(* IEC 61131-3 sources: plc-vscode/tests/st/all/trust-platform/crates/trust-runtime/tests/fixtures/ci/green/src, 1 file *)

(* ---- main.st ---- *)
PROGRAM Main
VAR
    Count : INT := 0;
END_VAR

Count := Count + 1;
END_PROGRAM
